FUNCTION_BLOCK Controle_PID_HMI (* Service Interface Function Block Type *)
  (* Standard: 61499-2 *)
  (* Version 1.0, 21/10/2026, Hidryco, Hidryco, IHM do Controle_PID *)
  PACKAGE Hidryco.HidrycoLib;
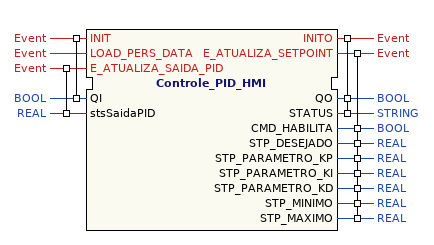
  EVENT_INPUT
    INIT WITH QI;
    LOAD_PERS_DATA; (* Reenvia os parametros persistentes *)
    E_ATUALIZA_SAIDA_PID WITH stsSaidaPID; (* Status do processo *)
  END_EVENT
  EVENT_OUTPUT
    INITO WITH QO, STATUS;
    E_ATUALIZA_SETPOINT WITH CMD_HABILITA, STP_DESEJADO, STP_PARAMETRO_KP, STP_PARAMETRO_KI, STP_PARAMETRO_KD, STP_MAXIMO, STP_MINIMO; (* Ajustes (IHM/OPC UA e LOAD_PERS_DATA) *)
  END_EVENT
  VAR_INPUT
    QI : BOOL;
    stsSaidaPID : REAL; (* Saida do PID (%) *)
  END_VAR
  VAR_OUTPUT
    QO : BOOL; (* Event Output Qualifier *)
    STATUS : STRING; (* Service Status *)
    CMD_HABILITA : BOOL; (* PID habilitado *)
    STP_DESEJADO : REAL; (* Valor desejado *)
    STP_PARAMETRO_KP : REAL; (* Ganho (Kp) *)
    STP_PARAMETRO_KI : REAL; (* Tempo integral (s) *)
    STP_PARAMETRO_KD : REAL; (* Tempo derivativo (s) *)
    STP_MINIMO : REAL; (* Saída mínima *)
    STP_MAXIMO : REAL; (* Saída máxima *)
  END_VAR
  SERVICE /
    SEQUENCE 
    END_SEQUENCE
  END_SERVICE
END_FUNCTION_BLOCK
